// TwinCAT 3 PLC project master
// ProgramVersion: 3.1.4026.27
// libraries:
//   Tc2_Standard, * (Beckhoff Automation GmbH)
//   Tc2_System, * (Beckhoff Automation GmbH)
//   Tc2_Utilities, * (Beckhoff Automation GmbH)
//   TcOtlp, * (S&E Engineering)
// project tree:
//   DUTs/ ST_SkidCommand.TcDUT, ST_SkidStatus.TcDUT
//   POUs/ FB_SkidClient.TcPOU
//   / GVL.TcGVL, MAIN.TcPOU, PlcTask.TcTTO
// real-time tasks:
//   TASK PlcTask: cycle T#10ms, priority 20, ADS port 350
//   TASK PlcTask1: cycle T#10ms, priority 21, ADS port 351
//   TASK PlcTask2: cycle T#10ms, priority 22, ADS port 352
//   TASK PlcTask3: cycle T#10ms, priority 23, ADS port 353

CONFIGURATION master
    RESOURCE PLC ON TwinCAT3
        TASK PlcTask(INTERVAL := T#10ms, PRIORITY := 20);
        PROGRAM MAIN WITH PlcTask : MAIN;
    END_RESOURCE
END_CONFIGURATION

// ---- DUTs/ST_SkidCommand.TcDUT
(*
	A stage command from the master to a pump skid, written to the skid's GVL.command in one ADS
	write so the carrier never arrives beside a stale command. The skid acts on a new sequence.
	Keep this identical to ST_SkidCommand in every skid project: ADS copies it byte for byte.
*)
TYPE ST_SkidCommand :
STRUCT
	sequence: UDINT;  // the master increments this for each command
	stageUp: BOOL;  // TRUE to stage up, FALSE to stage down
	flowRate: REAL;  // GPM
	carrier: ST_TraceContextCarrier;  // the master's client span, so the skid's spans join its trace
END_STRUCT
END_TYPE

// ---- DUTs/ST_SkidStatus.TcDUT
(*
	A pump skid's status, read by the master from the skid's GVL.status over ADS. A command has
	settled when sequence matches the command's and busy is clear.
	Keep this identical to ST_SkidStatus in every skid project: ADS copies it byte for byte.
*)
TYPE ST_SkidStatus :
STRUCT
	sequence: UDINT;  // the last command the skid accepted
	busy: BOOL;  // staging up or down, until the skid's staging span has ended
	running: BOOL;  // staged up
	faulted: BOOL;  // the last command ended in a fault
	faultText: STRING(80);  // why, when faulted
	flowRate: REAL;  // GPM
END_STRUCT
END_TYPE

// ---- GVL.TcGVL
{attribute 'qualified_only'}
VAR_GLOBAL
	// global logger provider
	resource: FB_Resource(schemaUrl:='');
	loggerProvider: FB_LoggerProvider(resource:=resource);
	
	// global tracer provider
	sampler: FB_Sampler_AlwaysOn();
	idGenerator: FB_IdGenerator(nTraceIds:=5, nSpanIds:=5);
	tracerProvider: FB_TracerProvider(resource:=resource, idGenerator:=idGenerator, sampler:=sampler);
END_VAR

// ---- MAIN.TcPOU
PROGRAM MAIN
VAR
	// logging config, note that loggers are oriented on a per entity (device) basis.
	staging: FB_InstrumentationScope(name:='staging', version:='0.0.0a', schemaUrl:='');
	masterLogger: FB_Logger(provider:=GVL.loggerProvider, scope:=staging);
	logExporter: FB_LogRecordExporter_HTTP('http://192.168.97.55:4318/v1/logs', TRUE);
	logBatchProcessor: FB_LogRecordProcessor_Batch(maxQueueSize:=500, scheduledDelayMillis:=1500,
												maxExportBatchSize:=500, exporter:=logExporter);

	// tracing config, note that tracers are oriented per service basis.
	tracer: FB_Tracer(scope:=staging, provider:=GVL.tracerProvider);
	spanExporter: FB_SpanExporter_HTTP('http://192.168.97.55:4318/v1/traces', TRUE);
	spanBatchProcessor: FB_SpanProcessor_Batch(maxQueueSize:=500, scheduledDelayMillis:=1500,
										   maxExportBatchSize:=500, exporter:=spanExporter);

	// the pump skids, each with one chiller; the name is the skid's service.name and the port its PLC's ADS port
	skid1: FB_SkidClient(tracer:=tracer, logger:=masterLogger, name:='pumpskid1', port:=852);
	skid2: FB_SkidClient(tracer:=tracer, logger:=masterLogger, name:='pumpskid2', port:=853);
	skid3: FB_SkidClient(tracer:=tracer, logger:=masterLogger, name:='pumpskid3', port:=854);

	// initialization setup
	firstScan: BOOL := TRUE;
	startupTimer: TON := (PT:=T#3S);  // lets the skid clients connect before the first staging decision

	// lead/lag/standby configuration
	{attribute 'OPC.UA.DA' := '1'}
	priority: ARRAY [0..2] OF USINT := [1, 2, 3];  // skid numbers, lead first
	{attribute 'OPC.UA.DA' := '1'}
	reqCount: USINT := 0;  // chillers required (in a real situation this would likely come from SCADA)
	{attribute 'OPC.UA.DA' := '1'}
	skidFlowRate: REAL := 700;  // GPM commanded to each skid that stages up

	// staging
	{attribute 'OPC.UA.DA' := '1'}
	runningCount: USINT;
	stagingState: USINT;
	stagingUp: BOOL;  // the direction of the sequence in progress
	attempted: ARRAY [1..3] OF BOOL;  // skids already commanded in this sequence, by skid number
	activeSkid: USINT;  // the skid whose command is in flight, 0 when none
	pStagingSpan: POINTER TO FB_Span;  // encloses every skid command of one sequence
	sequenceFailed: BOOL;  // the last sequence ran out of skids before reaching reqCount
	failedReqCount: USINT;  // the reqCount it failed on; a new reqCount retries at once
	retryTimer: TON := (PT:=T#30S);  // otherwise a failed sequence is retried after this
	skid: REFERENCE TO FB_SkidClient;
	candidate: USINT;
	skidNumber: USINT;
	i: USINT;
END_VAR

IF firstScan THEN
	GVL.resource.attributes
		.setStringAttribute('service.name', 'master_controller');
END_IF

// run the logger every tick
GVL.loggerProvider
	.stageProcessor(logBatchProcessor)
	.tick();

// run the tracer every tick
GVL.tracerProvider
	.stageProcessor(spanBatchProcessor)
	.tick();

// talk to the skids every tick
skid1();
skid2();
skid3();

runningCount := BOOL_TO_USINT(skid1.running) + BOOL_TO_USINT(skid2.running) + BOOL_TO_USINT(skid3.running);

startupTimer(IN:=TRUE);
retryTimer(IN:=stagingState = 0 AND sequenceFailed);

// perform the stage up or down to the desired number of chillers
CASE stagingState OF
	0: // settled: start a sequence when the running count differs from the required count
		IF startupTimer.Q AND runningCount <> reqCount
			AND (NOT sequenceFailed OR retryTimer.Q OR reqCount <> failedReqCount)
		THEN
			sequenceFailed := FALSE;
			stagingUp := reqCount > runningCount;
			MEMSET(ADR(attempted), 0, SIZEOF(attempted));
			tracer
				.startSpan(SEL(stagingUp, 'master.staging.stage_down', 'master.staging.stage_up'))
				.setNumberAttribute('chillers.required', reqCount)
				.setNumberAttribute('chillers.running', runningCount)
				.build(pStagingSpan);
			masterLogger
				.startLogRecord(E_SeverityNumber.INFO)
				.setBody(SEL(stagingUp, 'staging chillers down', 'staging chillers up'))
				.setNumberAttribute('chillers.required', reqCount)
				.setNumberAttribute('chillers.running', runningCount)
				.setTraceContextFromSpan(pStagingSpan)
				.emit();
			stagingState := 10;
		END_IF

	10: // command the next skid, or finish once enough are running
		IF runningCount = reqCount OR stagingUp <> (reqCount > runningCount) THEN
			// reached; or reqCount moved past the running count, and a new sequence starts from state 0
			tracer.setSpanStatusOk(pStagingSpan);
			tracer.endSpan(pStagingSpan);
			stagingState := 0;
		ELSE
			// stage up in priority order and down in reverse, so the lead skid runs longest
			candidate := 0;
			FOR i := 0 TO 2 DO
				skidNumber := priority[SEL(stagingUp, 2 - i, i)];
				skid REF= _skid(skidNumber);
				IF candidate = 0 AND __ISVALIDREF(skid) AND_THEN NOT attempted[skidNumber] AND skid.running <> stagingUp THEN
					candidate := skidNumber;
				END_IF
			END_FOR

			IF candidate = 0 THEN
				// every skid has been tried
				tracer.setSpanStatusError(pStagingSpan, SEL(stagingUp,
					'no running skid could be stopped',
					'not enough skids could be started'));
				masterLogger
					.startLogRecord(E_SeverityNumber.ERROR)
					.setBody(SEL(stagingUp,
						'staging down failed, no running skid could be stopped',
						'staging up failed, not enough skids could be started'))
					.setNumberAttribute('chillers.required', reqCount)
					.setNumberAttribute('chillers.running', runningCount)
					.setTraceContextFromSpan(pStagingSpan)
					.emit();
				tracer.endSpan(pStagingSpan);
				sequenceFailed := TRUE;
				failedReqCount := reqCount;
				stagingState := 0;
			ELSE
				attempted[candidate] := TRUE;
				skid REF= _skid(candidate);
				IF skid.command(stageUp:=stagingUp, flowRate:=skidFlowRate, pParentSpan:=pStagingSpan) THEN
					activeSkid := candidate;
					stagingState := 20;
				END_IF
			END_IF
		END_IF

	20: // wait for the skid to settle; after a failure, state 10 moves on to the next skid
		skid REF= _skid(activeSkid);
		IF NOT __ISVALIDREF(skid) OR_ELSE skid.commandDone THEN
			activeSkid := 0;
			stagingState := 10;
		END_IF
END_CASE

firstScan := FALSE;

(* The skid client with the given number, or an invalid reference for any other number. *)
METHOD _skid : REFERENCE TO FB_SkidClient
VAR_INPUT
	number: USINT;
END_VAR
CASE number OF
	1: _skid REF= skid1;
	2: _skid REF= skid2;
	3: _skid REF= skid3;
END_CASE
END_METHOD

END_PROGRAM

// ---- POUs/FB_SkidClient.TcPOU
(*
	The master's side of one pump skid. It polls the skid's GVL.status over ADS and writes stage
	commands to its GVL.command.

	Each command runs inside a CLIENT span whose context travels with the command in an
	ST_TraceContextCarrier. The skid extracts it and parents its SERVER staging span on it, so
	the skid's spans sit inside this one and the service graph shows master -> skid. The client
	span ends only once the skid reports it has settled, which is after the skid's staging span
	has ended, so the skid's spans are fully enclosed.

	Call the block every cycle. command starts a command; commandDone and commandOk report how it
	ended. A skid that cannot be reached fails its command at once, with an error span and log,
	so the caller can move on to the next skid.
*)
FUNCTION_BLOCK FB_SkidClient
VAR_INPUT
	netId: T_AmsNetId := '';  // '' is this machine
END_VAR
VAR_OUTPUT
	online: BOOL;  // both handles granted and the last status read succeeded
	status: ST_SkidStatus;  // the last status read from the skid
	running: BOOL;  // online and staged up
	commandBusy: BOOL;  // a command is in flight
	commandDone: BOOL;  // the last command has ended; stays set until the next command
	commandOk: BOOL;  // the last command left the skid in the commanded state
	adsErrorId: UDINT;  // the last ADS error, 0 once a connection succeeds
END_VAR
VAR CONSTANT
	ADSIGRP_SYM_HNDBYNAME: UDINT := 16#F003;  // get a handle for a symbol name
	ADSIGRP_SYM_VALBYHND: UDINT := 16#F005;  // read or write a symbol through its handle
	ADSIGRP_SYM_RELEASEHND: UDINT := 16#F006;  // release a handle
	ADS_TIMEOUT: TIME := T#1S;  // each ADS request gives up after this
	POLL_PERIOD: TIME := T#200MS;
	RECONNECT_DELAY: TIME := T#5S;
	COMMAND_TIMEOUT: TIME := T#3M;  // longer than the slowest simulated stage up
END_VAR
VAR
	_tracer: REFERENCE TO FB_Tracer;
	_logger: REFERENCE TO FB_Logger;
	_name: STRING;  // the skid's service.name, used as peer.service
	_port: UINT;  // the skid PLC's ADS port

	_commandSymbol: STRING := 'GVL.command';
	_statusSymbol: STRING := 'GVL.status';
	_command: ST_SkidCommand;  // stays put while a write is in flight
	_received: ST_SkidStatus;  // reads land here, so status only changes on a good read
	_commandHandle: UDINT;
	_statusHandle: UDINT;
	_hasCommandHandle: BOOL;
	_hasStatusHandle: BOOL;

	_getHandle: ADSRDWRT;
	_read: ADSREAD;
	_write: ADSWRITE;
	_releaseHandle: ADSWRITE;
	_state: USINT;
	_pollTimer: TON;
	_reconnectTimer: TON;
	_commandTimer: TON;

	_sendPending: BOOL;  // command was called and the write has not been issued yet
	_awaitingSkid: BOOL;  // the write landed; waiting for the skid to settle
	_pSpan: POINTER TO FB_Span;  // the CLIENT span of the command in flight; owned here until it ends
END_VAR

_pollTimer(IN:=NOT _pollTimer.Q, PT:=POLL_PERIOD);
_reconnectTimer(IN:=_state = 90, PT:=RECONNECT_DELAY);
_commandTimer(IN:=_awaitingSkid, PT:=COMMAND_TIMEOUT);

IF _commandTimer.Q THEN
	THIS^._finishCommand(ok:=FALSE, message:=CONCAT(_name, ' did not settle before the command timed out'));
END_IF

CASE _state OF
	0: // ask the skid for a handle to its command symbol
		_getHandle(
			NETID:=netId,
			PORT:=_port,
			IDXGRP:=ADSIGRP_SYM_HNDBYNAME,
			IDXOFFS:=0,
			WRITELEN:=TO_UDINT(LEN(_commandSymbol)),
			READLEN:=SIZEOF(_commandHandle),
			SRCADDR:=ADR(_commandSymbol),
			DESTADDR:=ADR(_commandHandle),
			WRTRD:=TRUE,
			TMOUT:=ADS_TIMEOUT);
		_state := 10;

	10: // wait for the command handle, then ask for the status handle
		_getHandle(WRTRD:=FALSE);
		IF NOT _getHandle.BUSY THEN
			IF _getHandle.ERR THEN
				THIS^._goOffline(errorId:=_getHandle.ERRID);
			ELSE
				_hasCommandHandle := TRUE;
				_getHandle(
					NETID:=netId,
					PORT:=_port,
					IDXGRP:=ADSIGRP_SYM_HNDBYNAME,
					IDXOFFS:=0,
					WRITELEN:=TO_UDINT(LEN(_statusSymbol)),
					READLEN:=SIZEOF(_statusHandle),
					SRCADDR:=ADR(_statusSymbol),
					DESTADDR:=ADR(_statusHandle),
					WRTRD:=TRUE,
					TMOUT:=ADS_TIMEOUT);
				_state := 20;
			END_IF
		END_IF

	20: // wait for the status handle, then read the status once before going online
		_getHandle(WRTRD:=FALSE);
		IF NOT _getHandle.BUSY THEN
			IF _getHandle.ERR THEN
				THIS^._goOffline(errorId:=_getHandle.ERRID);
			ELSE
				_hasStatusHandle := TRUE;
				THIS^._readStatus();
				_state := 30;
			END_IF
		END_IF

	30: // the first read: continue from the skid's sequence, so a restarted master never repeats an old one
		_read(READ:=FALSE);
		IF NOT _read.BUSY THEN
			IF _read.ERR THEN
				THIS^._goOffline(errorId:=_read.ERRID);
			ELSE
				status := _received;
				_command.sequence := status.sequence;
				adsErrorId := 0;
				online := TRUE;
				_state := 40;
			END_IF
		END_IF

	40: // online and idle: a pending command goes out before the next poll
		IF _sendPending THEN
			_sendPending := FALSE;
			// the command and its carrier in one write, so the skid never sees one without the other
			_write(
				NETID:=netId,
				PORT:=_port,
				IDXGRP:=ADSIGRP_SYM_VALBYHND,
				IDXOFFS:=_commandHandle,
				LEN:=SIZEOF(_command),
				SRCADDR:=ADR(_command),
				WRITE:=TRUE,
				TMOUT:=ADS_TIMEOUT);
			_state := 50;
		ELSIF _pollTimer.Q THEN
			THIS^._readStatus();
			_state := 60;
		END_IF

	50: // wait for the command to land
		_write(WRITE:=FALSE);
		IF NOT _write.BUSY THEN
			IF _write.ERR THEN
				THIS^._goOffline(errorId:=_write.ERRID);
			ELSE
				_awaitingSkid := TRUE;
				_state := 40;
			END_IF
		END_IF

	60: // wait for the status; a command has settled once the skid has accepted it and is no longer busy
		_read(READ:=FALSE);
		IF NOT _read.BUSY THEN
			IF _read.ERR THEN
				THIS^._goOffline(errorId:=_read.ERRID);
			ELSE
				status := _received;
				IF _awaitingSkid AND status.sequence = _command.sequence AND NOT status.busy THEN
					IF status.running = _command.stageUp THEN
						THIS^._finishCommand(ok:=TRUE, message:=CONCAT(_name, SEL(_command.stageUp, ' staged down', ' staged up')));
					ELSIF status.faulted THEN
						THIS^._finishCommand(
							ok:=FALSE,
							message:=CONCAT(CONCAT(_name, SEL(_command.stageUp, ' failed to stage down: ', ' failed to stage up: ')), status.faultText));
					ELSE
						THIS^._finishCommand(ok:=FALSE, message:=CONCAT(_name, ' settled without reaching the commanded state'));
					END_IF
				END_IF
				_state := 40;
			END_IF
		END_IF

	70: // release the command handle, if one was granted
		IF _hasCommandHandle THEN
			_releaseHandle(
				NETID:=netId,
				PORT:=_port,
				IDXGRP:=ADSIGRP_SYM_RELEASEHND,
				IDXOFFS:=0,
				LEN:=SIZEOF(_commandHandle),
				SRCADDR:=ADR(_commandHandle),
				WRITE:=TRUE,
				TMOUT:=ADS_TIMEOUT);
			_state := 75;
		ELSE
			_state := 80;
		END_IF

	75: // a failed release only leaves a handle on a skid that has gone away
		_releaseHandle(WRITE:=FALSE);
		IF NOT _releaseHandle.BUSY THEN
			_hasCommandHandle := FALSE;
			_state := 80;
		END_IF

	80: // release the status handle, if one was granted
		IF _hasStatusHandle THEN
			_releaseHandle(
				NETID:=netId,
				PORT:=_port,
				IDXGRP:=ADSIGRP_SYM_RELEASEHND,
				IDXOFFS:=0,
				LEN:=SIZEOF(_statusHandle),
				SRCADDR:=ADR(_statusHandle),
				WRITE:=TRUE,
				TMOUT:=ADS_TIMEOUT);
			_state := 85;
		ELSE
			_state := 90;
		END_IF

	85:
		_releaseHandle(WRITE:=FALSE);
		IF NOT _releaseHandle.BUSY THEN
			_hasStatusHandle := FALSE;
			_state := 90;
		END_IF

	90: // offline: wait, then connect again
		IF _reconnectTimer.Q THEN
			_state := 0;
		END_IF
END_CASE

running := online AND status.running;

(*
	Starts a stage command inside a new CLIENT span, a child of pParentSpan when one is given.
	The span's context is injected into the command's carrier for the skid to extract. Returns
	FALSE, and changes nothing, while a command is already in flight. A skid that is not online
	fails the command at once, so commandDone is already set when this returns.
*)
METHOD command : BOOL
VAR_INPUT
	stageUp: BOOL;  // TRUE to stage up, FALSE to stage down
	flowRate: REAL;  // GPM
	pParentSpan: POINTER TO FB_Span;  // borrowed for the call: the client span becomes its child
END_VAR
VAR
	_pContext: POINTER TO FB_SpanContext;
END_VAR
command := FALSE;

IF commandBusy THEN
	RETURN;
END_IF

commandBusy := TRUE;
commandDone := FALSE;
commandOk := FALSE;

_tracer
	.startSpan(name:=SEL(stageUp, 'skid.command.stage_down', 'skid.command.stage_up'), kind:=E_SpanKind.SPAN_KIND_CLIENT)
	.setStringAttribute('peer.service', _name)
	.setStringAttribute('rpc.system', 'ads')
	.setNumberAttribute('server.port', _port)
	.setNumberAttribute('flow.target', flowRate);
IF pParentSpan <> 0 THEN
	_tracer.setParentUsingSpan(pParentSpan);
END_IF
_tracer.build(pDest:=_pSpan);

// without a span the carrier goes out empty, and the skid starts its own trace
MEMSET(ADR(_command.carrier), 0, SIZEOF(_command.carrier));
IF _tracer.getSpanContext(pDest:=_pContext, pSpan:=_pSpan) THEN
	TraceContextPropagator.inject(pContext:=_pContext, carrier:=_command.carrier);
	_pContext^.delete(pSelf:=_pContext);
END_IF

_command.sequence := _command.sequence + 1;
_command.stageUp := stageUp;
_command.flowRate := flowRate;

IF online THEN
	_sendPending := TRUE;
ELSIF adsErrorId <> 0 THEN
	THIS^._finishCommand(ok:=FALSE, message:=CONCAT(CONCAT(_name, ' is unreachable, ADS error '), UDINT_TO_STRING(adsErrorId)));
ELSE
	THIS^._finishCommand(ok:=FALSE, message:=CONCAT(_name, ' is not connected yet'));
END_IF

command := TRUE;
END_METHOD

METHOD FB_Exit : BOOL
VAR_INPUT
	bInCopyCode: BOOL;  // TRUE: the exit method is called in order to leave the instance which will be copied afterwards (online change).
END_VAR
// during an online change the copied instance keeps the span
IF NOT bInCopyCode THEN
	_tracer.discardSpan(pSpan:=_pSpan);
END_IF
END_METHOD

METHOD FB_Init : BOOL
VAR_INPUT
	bInitRetains: BOOL;  // TRUE: the retain variables are initialized (reset warm / reset cold)
	bInCopyCode: BOOL;  // TRUE: the instance will be copied to the copy code afterward (online change)
	tracer: REFERENCE TO FB_Tracer;  // starts and ends the command spans
	logger: REFERENCE TO FB_Logger;  // logs how each command ended
	name: STRING;  // the skid's service.name, used as peer.service
	port: UINT;  // the skid PLC's ADS port
END_VAR
THIS^._tracer REF= tracer;
THIS^._logger REF= logger;
THIS^._name := name;
THIS^._port := port;
END_METHOD

(* Ends the command in flight: sets its span's status, logs the outcome in the span, and ends the span. *)
METHOD _finishCommand
VAR_INPUT
	ok: BOOL;
	message: T_MaxString;
END_VAR
commandBusy := FALSE;
commandDone := TRUE;
commandOk := ok;
_sendPending := FALSE;
_awaitingSkid := FALSE;

IF ok THEN
	_tracer.setSpanStatusOk(pSpan:=_pSpan);
	_logger
		.startLogRecord(E_SeverityNumber.INFO)
		.setBody(message)
		.setStringAttribute('peer.service', _name)
		.setTraceContextFromSpan(_pSpan)
		.emit();
ELSE
	_tracer.setSpanStatusError(pSpan:=_pSpan, message:=message);
	_logger
		.startLogRecord(E_SeverityNumber.ERROR)
		.setBody(message)
		.setStringAttribute('peer.service', _name)
		.setTraceContextFromSpan(_pSpan)
		.emit();
END_IF

_tracer.endSpan(pSpan:=_pSpan);
END_METHOD

(* Drops the connection after an ADS error: fails any command in flight, then releases the handles and waits to reconnect. *)
METHOD _goOffline
VAR_INPUT
	errorId: UDINT;
END_VAR
online := FALSE;
adsErrorId := errorId;

IF commandBusy THEN
	THIS^._finishCommand(ok:=FALSE, message:=CONCAT(CONCAT(_name, ' is unreachable, ADS error '), UDINT_TO_STRING(errorId)));
END_IF

_state := 70;
END_METHOD

(* Starts a read of the skid's status into _received. *)
METHOD _readStatus
_read(
	NETID:=netId,
	PORT:=_port,
	IDXGRP:=ADSIGRP_SYM_VALBYHND,
	IDXOFFS:=_statusHandle,
	LEN:=SIZEOF(_received),
	DESTADDR:=ADR(_received),
	READ:=TRUE,
	TMOUT:=ADS_TIMEOUT);
END_METHOD

END_FUNCTION_BLOCK
